(* IEC 61131-3 sources: llm-plc-st-eval/data/raw/claude-sonnet-4-6/I6/few_shot, 3 files *)

(* ---- ejec_1.st ---- *)
```pascal
FUNCTION_BLOCK FB_Temperatura
VAR_INPUT
    rawTemp : INT; (* Valor crudo del sensor: 0..27648 -> 0.0..100.0 °C *)
END_VAR
VAR_OUTPUT
    tempC     : REAL; (* Temperatura calculada en grados Celsius *)
    enfriador : BOOL; (* Salida del enfriador *)
    almSensor : BOOL; (* Alarma de sensor fuera de rango *)
END_VAR

(* Verificar rango valido del sensor *)
IF rawTemp < 0 OR rawTemp > 27648 THEN
    almSensor := TRUE;
    enfriador := FALSE; (* Apagar enfriador por seguridad ante fallo *)
ELSE
    almSensor := FALSE;

    (* Escalar valor crudo a grados Celsius: tempC = rawTemp * 100.0 / 27648.0 *)
    tempC := INT_TO_REAL(rawTemp) * 100.0 / 27648.0;

    (* Control con histeresis: ON >= 80.0, OFF <= 75.0, entre ambos conserva estado *)
    IF tempC >= 80.0 THEN
        enfriador := TRUE;  (* Activar enfriador al superar umbral alto *)
    ELSIF tempC <= 75.0 THEN
        enfriador := FALSE; (* Desactivar enfriador al bajar del umbral bajo *)
    (* Entre 75.0 y 80.0 exclusivo: enfriador mantiene su estado anterior *)
    END_IF;
END_IF;

END_FUNCTION_BLOCK
```

(* ---- ejec_2.st ---- *)
```pascal
FUNCTION_BLOCK FB_Temperatura
VAR_INPUT
    rawTemp : INT; (* Valor crudo del sensor: 0..27648 -> 0.0..100.0 °C *)
END_VAR
VAR_OUTPUT
    tempC     : REAL; (* Temperatura calculada en grados Celsius *)
    enfriador : BOOL; (* Salida del enfriador *)
    almSensor : BOOL; (* Alarma de sensor fuera de rango *)
END_VAR
VAR CONSTANT
    RAW_MIN  : INT  := 0;       (* Valor crudo minimo valido *)
    RAW_MAX  : INT  := 27648;   (* Valor crudo maximo valido *)
    TEMP_MAX : REAL := 100.0;   (* Temperatura maxima de escala *)
    HIS_ON   : REAL := 80.0;    (* Umbral de activacion del enfriador *)
    HIS_OFF  : REAL := 75.0;    (* Umbral de desactivacion del enfriador *)
END_VAR

(* --- Verificacion de rango del sensor --- *)
IF rawTemp < RAW_MIN OR rawTemp > RAW_MAX THEN
    almSensor := TRUE;   (* Fuera de rango: activa alarma *)
    enfriador := FALSE;  (* Apaga el enfriador por seguridad *)
    tempC     := 0.0;    (* Valor de temperatura indefinido *)
ELSE
    almSensor := FALSE;

    (* --- Conversion lineal: rawTemp -> grados Celsius --- *)
    (* tempC = (rawTemp / 27648) * 100.0                   *)
    tempC := (INT_TO_REAL(rawTemp) / INT_TO_REAL(RAW_MAX)) * TEMP_MAX;

    (* --- Control con histeresis --- *)
    IF tempC >= HIS_ON THEN
        enfriador := TRUE;   (* Supera umbral alto: enciende enfriador *)
    ELSIF tempC <= HIS_OFF THEN
        enfriador := FALSE;  (* Baja del umbral bajo: apaga enfriador *)
    (* Entre 75.0 y 80.0: conserva el estado anterior (histeresis) *)
    END_IF;
END_IF;

END_FUNCTION_BLOCK
```

(* ---- ejec_3.st ---- *)
```pascal
FUNCTION_BLOCK FB_Temperatura
VAR_INPUT
    rawTemp : INT; (* Valor crudo del sensor: 0..27648 -> 0.0..100.0 °C *)
END_VAR
VAR_OUTPUT
    tempC     : REAL; (* Temperatura calculada en grados Celsius *)
    enfriador : BOOL; (* Salida del enfriador *)
    almSensor : BOOL; (* Alarma de sensor fuera de rango *)
END_VAR

(* Verificar rango valido del sensor *)
IF rawTemp < 0 OR rawTemp > 27648 THEN
    almSensor := TRUE;
    enfriador := FALSE; (* Enfriador desactivado por fallo de sensor *)
ELSE
    almSensor := FALSE;

    (* Conversion lineal: tempC = rawTemp * 100.0 / 27648.0 *)
    tempC := INT_TO_REAL(rawTemp) * 100.0 / 27648.0;

    (* Control con histeresis: enciende >= 80.0, apaga <= 75.0 *)
    IF tempC >= 80.0 THEN
        enfriador := TRUE;
    ELSIF tempC <= 75.0 THEN
        enfriador := FALSE;
    (* Entre 75.0 y 80.0 exclusivo: conserva el estado anterior *)
    END_IF;
END_IF;

END_FUNCTION_BLOCK
```
